// TIA Portal V17 export
FUNCTION "Mini_FC" : Void   // FC1, LAD
   VAR_TEMP
      Tmp : Bool;
   END_VAR
BEGIN

REGION Network 1: Пуск двигателя
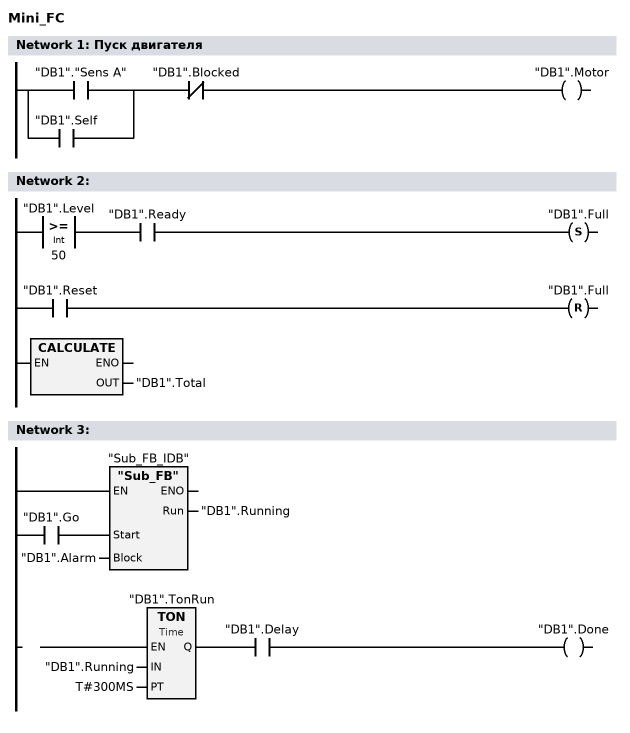
   RUNG wire#powerrail
      Contact( "DB1"."Sens A" )
      wire#w1
      I_Contact( "DB1".Blocked )
      Coil( "DB1".Motor )
   END_RUNG
   RUNG wire#powerrail
      Contact( "DB1".Self )
   END_RUNG wire#w1
   // the same network as SCL:
   "DB1".Motor := ("DB1"."Sens A" OR "DB1".Self) AND NOT "DB1".Blocked;
END_REGION

REGION Network 2
   RUNG wire#powerrail
      { S7_Templates := "SrcType := Int" } GE_Contact(in1 := "DB1".Level, in2 := 50)
      Contact( "DB1".Ready )
      S_Coil( "DB1".Full )
   END_RUNG
   RUNG wire#powerrail
      Contact( "DB1".Reset )
      R_Coil( "DB1".Full )
   END_RUNG
   RUNG wire#powerrail
      { S7_GenerateENO := "TRUE" } Calculate(out => "DB1".Total)
   END_RUNG
   // the same network as SCL:
   // no SCL statement known for Calc: written as a call
   IF ("DB1".Level >= 50) AND "DB1".Ready THEN "DB1".Full := TRUE; END_IF;
   IF "DB1".Reset THEN "DB1".Full := FALSE; END_IF;
   Calc(out => "DB1".Total);
END_REGION

REGION Network 3
   "Sub_FB_IDB"(Start := "DB1".Go, Block := "DB1".Alarm, Run => "DB1".Running);   // "Sub_FB"
   "DB1".TonRun.TON(IN := "DB1".Running, PT := T#300MS);
   "DB1".Done := "DB1".TonRun.Q AND "DB1".Delay;
END_REGION
END_FUNCTION
